Fanuc KAREL source: kb00123.KL

-- PROVISIONAL review KL for V1013-1; original PC SHA256 e094456801df9577bc554bcbdfd31a0f0d1bb33582b5694cdc6aa6b9c7718ff8
-- Incomplete behavior may be omitted. Consult companion uncertainty JSON. Do not deploy.
PROGRAM KB00123
%NOLOCKGROUP
BEGIN
  -- UNRESOLVED_PC offsets 5-14; opcodes 3F,75
  -- UNRESOLVED_PC offsets 19-26; opcodes 9D,23
  -- UNRESOLVED_PC offsets 31-49; opcodes 27,22,2A,22,31
  -- UNRESOLVED_PC offsets 54-58; opcodes 7F
END KB00123
